// TIA Portal V21 export
DATA_BLOCK "IDB_Doser"   // DB6
// stored: InstanceOfName Dosing.FB_Doser, InstanceOfType FB, Namespace Dosing
"Dosing.FB_Doser"
   // VAR_INPUT
   //    Start : Bool;
   //    Stop : Bool;
   // END_VAR
   // VAR_OUTPUT
   //    Dosing : Bool;
   //    Done : Bool;
   // END_VAR
   // VAR
   //    Filler { S7_SetPoint := 'True'} : "Filling.FB_Filler";
   //    Recipe { S7_SetPoint := 'True'} : "Filling.UDT_FillRecipe";
   // END_VAR
BEGIN
END_DATA_BLOCK
